FUNCTION_BLOCK TcoMessengerTests EXTENDS TcoCore.TcoObject
VAR
	_category : TcoCore.eMessageCategory;
	_minLevel : TcoCore.eMessageCategory;
	_messageDigestMethod : TcoCore.eMessageDigestMethod;
	_messageLoggingMethod : TcoCore.eMessengerLogMethod;
END_VAR

VAR
	_BOOL			: BOOL 				 := TRUE;
	_BYTE			: BYTE				 := 1;
	_WORD			: WORD				 := 22;
	_DWORD			: DWORD				 := 333;
	_LWORD			: LWORD				 := 4444;
	_SINT			: SINT				 := 12;
	_USINT			: USINT				 := 13;
	_INT			: INT				 := 14; 
	_UINT			: UINT				 := 55;
	_DINT			: DINT				 := 66;
	_UDINT			: UDINT				 := 77;
	_LINT			: LINT				 := 88;
	_ULINT			: ULINT				 := 99;
	_LTIME			: LTIME				 :=	LTIME#551US615NS; 
	_Real 			: REAL				 := 99.9;
	_LReal			: LREAL				 :=	88.8;
	_DateAndTime 	: DATE_AND_TIME	 := DT#2106-02-06-06:28:15;
	_Date			: DATE				 := D#2106-02-06;
	_Time			: TIME				 := T#71582M47S295MS;
	_WString		: WSTRING			 := "W1";
	_TOD			: TOD				 := TOD#23:59:59.999;
	_String			: STRING			 :=	'S1';
END_VAR

{attribute 'TcRpcEnable'}
METHOD AppendAnys_1 : BOOL
VAR_INPUT
END_VAR
_messenger.Build().AppendAny(_BOOL		     )
                  .AppendAny(_BYTE		     )
                  .AppendAny(_WORD		     )
                  .AppendAny(_DWORD		     )
                  .AppendAny(_LWORD		     )
                  .AppendAny(_SINT		     )
                  .AppendAny(_USINT		     )
                  .AppendAny(_INT		     )
                  .AppendAny(_UINT		     )
                  .AppendAny(_DINT		     )
				  .AppendAny(_UDINT		     ).As().AsDebug();
END_METHOD

{attribute 'TcRpcEnable'}
METHOD AppendAnys_2 : BOOL
VAR_INPUT
END_VAR
_messenger.Build().AppendAny(_LINT		     )
				  .AppendAny(_ULINT		     )
				  .AppendAny(_LTIME		     )
                  .AppendAny(_Real 		     )
				  .AppendAny(_LReal		     )
				  .AppendAny(_DateAndTime    )
				  .AppendAny(_Date		     )  
                  .AppendAny(_Time		     )
				  .AppendAny(_WString	     )
				  .AppendAny(_TOD		     )
				  .AppendAny(_String		 ).As().AsDebug();
END_METHOD

{attribute 'TcRpcEnable'}
METHOD AsDebug : BOOL
VAR_INPUT
	TextMessage1 : STRING;
	TextMessage2 : STRING;
	Value : LREAL;
END_VAR
_messenger.Build().Append(TextMessage1).Append(TextMessage2).AppendAny(Value).As().AsDebug();
END_METHOD

{attribute 'TcRpcEnable'}
METHOD AsError : BOOL
VAR_INPUT
	TextMessage1 : STRING;
	TextMessage2 : STRING;
	Value : LREAL;
END_VAR
_messenger.Build().Append(TextMessage1).Append(TextMessage2).AppendAny(Value).As().AsError();
END_METHOD

{attribute 'TcRpcEnable'}
METHOD AsFatal : BOOL
VAR_INPUT
	TextMessage1 : STRING;
	TextMessage2 : STRING;
	Value : LREAL;
END_VAR
_messenger.Build().Append(TextMessage1).Append(TextMessage2).AppendAny(Value).As().AsFatal();
END_METHOD

{attribute 'TcRpcEnable'}
METHOD AsInfo : BOOL
VAR_INPUT
	TextMessage1 : STRING;
	TextMessage2 : STRING;
	Value : LREAL;
END_VAR
_messenger.Build().Append(TextMessage1).Append(TextMessage2).AppendAny(Value).As().AsInfo();
END_METHOD

{attribute 'TcRpcEnable'}
METHOD AsTrace : BOOL
VAR_INPUT
	TextMessage1 : STRING;
	TextMessage2 : STRING;
	Value : LREAL;
END_VAR
_messenger.Build().Append(TextMessage1).Append(TextMessage2).AppendAny(Value).As().AsTrace();
END_METHOD

{attribute 'TcRpcEnable'}
METHOD AsWarning : BOOL
VAR_INPUT
	TextMessage1 : STRING;
	TextMessage2 : STRING;
	Value : LREAL;
END_VAR
_messenger.Build().Append(TextMessage1).Append(TextMessage2).AppendAny(Value).As().AsWarning();
END_METHOD

{attribute 'TcRpcEnable'}
METHOD INTERNAL Catastrophic
VAR_INPUT	
	Message : STRING(255);
END_VAR
_messenger.Catastrophic(Message);
END_METHOD

{attribute 'TcRpcEnable'}
METHOD INTERNAL Critical
VAR_INPUT
	Message : STRING(255);
END_VAR
_messenger.Critical(Message);
END_METHOD

{attribute 'TcRpcEnable'}
METHOD INTERNAL Debug
VAR_INPUT
	Message : STRING(255);
END_VAR
_messenger.Debug(Message);
END_METHOD

{attribute 'TcRpcEnable'}
METHOD INTERNAL Error
VAR_INPUT
	Message : STRING(255);
END_VAR
_messenger.Error(Message);
END_METHOD

{attribute 'TcRpcEnable'}
METHOD INTERNAL Info
VAR_INPUT
	Message : STRING(255);
END_VAR
_messenger.Info(Message);
END_METHOD

{attribute 'TcRpcEnable'}
METHOD INTERNAL Notify
VAR_INPUT
	Message : STRING(255);
END_VAR
_messenger.Notify(Message);
END_METHOD

{attribute 'TcRpcEnable'}
METHOD OnCondition : BOOL
VAR_INPUT
	inCondition : BOOL;
	message : STRING;
END_VAR
_messenger.OnCondition(inCondition).Post(message, _category);
END_METHOD

{attribute 'TcRpcEnable'}
METHOD Pin : BOOL
VAR_INPUT
	inCondition : BOOL;
	message : STRING;
END_VAR
IF(inCondition)THEN
	_messenger.Post(message, _category).Pin();
ELSE
	_messenger.Post(message, _category);
END_IF;
END_METHOD

{attribute 'TcRpcEnable'}
METHOD Pinned : BOOL
Pinned := _messenger.Pinned;
END_METHOD

{attribute 'TcRpcEnable'}
METHOD INTERNAL Post 
VAR_INPUT	
	Message : STRING(255);	
END_VAR
_messenger.Post(Message, _category);
END_METHOD

{attribute 'TcRpcEnable'}
METHOD INTERNAL Programming
VAR_INPUT
	Message : STRING(255);
END_VAR
_messenger.Programming(Message);
END_METHOD

{attribute 'TcRpcEnable'}
METHOD INTERNAL Resume
Context.Environment.Messaging.Resume();
END_METHOD

{attribute 'TcRpcEnable'}
METHOD INTERNAL SetMessageDigestMethod
Context.Environment.Messaging.MessageDigestMethod := _messageDigestMethod;
END_METHOD

{attribute 'TcRpcEnable'}
METHOD INTERNAL SetMessageLoggingMethod
Context.Environment.Messaging.MessengerLoggingMethod := _messageLoggingMethod;
END_METHOD

{attribute 'TcRpcEnable'}
METHOD INTERNAL SetMinLevel
Context.Environment.Messaging.MinLevel := _minLevel;
END_METHOD

{attribute 'TcRpcEnable'}
METHOD INTERNAL Suspend
Context.Environment.Messaging.Suspend();
END_METHOD

{attribute 'TcRpcEnable'}
METHOD INTERNAL TimedOut
VAR_INPUT
	Message : STRING(255);
END_VAR
_messenger.Warning(Message);
END_METHOD

{attribute 'TcRpcEnable'}
METHOD INTERNAL Trace
VAR_INPUT
	Message : STRING(255);
END_VAR
_messenger.Trace(Message);
END_METHOD

{attribute 'TcRpcEnable'}
METHOD UnPin : BOOL
VAR_INPUT
	inCondition : BOOL;
	message : STRING;
END_VAR
_messenger.UnPin();
END_METHOD

{attribute 'TcRpcEnable'}
METHOD INTERNAL Warning
VAR_INPUT
	Message : STRING(255);
END_VAR
_messenger.Warning(Message);
END_METHOD

END_FUNCTION_BLOCK

(* stored: Version 1.1.0.1
   POU TcoMessengerTests: Id {d87e08d3-1876-01a7-16f8-c33755c3cedd}, SpecialFunc None
   Folder As: Id {8f4655ae-f441-09fd-2886-71c54526cb3c}
   Method AppendAnys_1: Id {75e9fff2-0d79-0c6b-1899-64e8e72ac807}
   Method AppendAnys_2: Id {cda3da18-b30b-0e91-1459-47c79d7fbf42}
   Method AsDebug: Id {28278033-884e-0754-16b7-a71ef9f36b70}
   Method AsError: Id {11de2039-508e-077a-3c59-04d05bc193fa}
   Method AsFatal: Id {3eebfd32-39af-088f-1125-85723e6f1daa}
   Method AsInfo: Id {0dd75bcc-a12d-0170-0caa-286251b11a98}
   Method AsTrace: Id {e5c2f330-7172-009a-258e-6e097bb33bef}
   Method AsWarning: Id {24d5dc4e-60b0-00a4-369e-a2d7751c346b}
   Method Catastrophic: Id {093578d4-4883-02db-1234-cd38a177e6a9}
   Method Critical: Id {cc04394e-ff89-0912-0edc-b599a0c7d07c}
   Method Debug: Id {d279de92-cd96-029d-39a9-f59f29b03fe7}
   Method Error: Id {8cdb9a84-d1f9-0d5c-21aa-e984960b0322}
   Method Info: Id {c925a1ca-2a19-0552-0bb5-9de32cfb972b}
   Method Notify: Id {32b9cbb6-6207-0f35-1241-0cd0d8f3e2c6}
   Method OnCondition: Id {e703b1c7-cb4e-0f53-157b-b659f402335a}
   Method Pin: Id {6f3b1ff2-ee84-08b3-3106-aabf05111047}
   Method Pinned: Id {b0bb481b-a0e8-0eda-3566-10e1585625b7}
   Method Post: Id {aa4eba68-8e3e-0790-14e4-37c20eb0fa3d}
   Method Programming: Id {ad9b3a9b-2e3a-01d3-03b2-0966d6f79bec}
   Method Resume: Id {82062340-d28d-08df-1727-1ea7f90e73d2}
   Method SetMessageDigestMethod: Id {f159a2ac-72e9-0d3d-2b2d-e8b8d72302e3}
   Method SetMessageLoggingMethod: Id {97fd978e-924e-0e25-274f-3c8a2c023916}
   Method SetMinLevel: Id {14062f88-3c36-0c8f-1769-35d9d0ae9a98}
   Method Suspend: Id {009042cd-d9d8-01ec-1e53-e01d1459f156}
   Method TimedOut: Id {df75203d-ff31-0992-037d-6d10558ac6d6}
   Method Trace: Id {02a9dc17-bef6-0f75-27b7-d7639e83bf18}
   Method UnPin: Id {19d9f139-709a-0227-3e03-cbb3323497b3}
   Method Warning: Id {032a7c5b-ea22-0043-0563-7ca4d7b308c3} *)
